(* IEC 61131-3 sources: plc-process-lib/tests/POUs/Helpers/FB_TestDeviceNoSuper, 1 file *)

(* ---- FB_TestDeviceNoSuper.decl.st ---- *)
// Назначение: наследник FB_TestDevice со своим телом без SUPER^: проверка во время выполнения,
//             что тело базы при вызове наследника само не выполняется (L1 контракта). Только для
//             тестов.
// Автор:      kr0nsch
// Версия:     0.1.0
// Документ:   docs/TESTING.md, раздел «Тестовое устройство»
FUNCTION_BLOCK FB_TestDeviceNoSuper EXTENDS FB_TestDevice
VAR
    uiOwnBodyCalls : UINT;       // сколько раз выполнено это тело
END_VAR
